(* IEC 61131-3 sources: trust-platform/examples/OSCAT/irrigation_sun_clock/non-oop/src, 1 file *)

(* ---- Configuration.st ---- *)
CONFIGURATION IrrigationSunClockClassicConfiguration
RESOURCE IrrigationSunClockClassic ON PLC
    TASK MainTask (INTERVAL := T#1s, PRIORITY := 1);
    PROGRAM Main WITH MainTask : Main;
END_RESOURCE
END_CONFIGURATION
